KUKA KRL program: DrillingPart.src

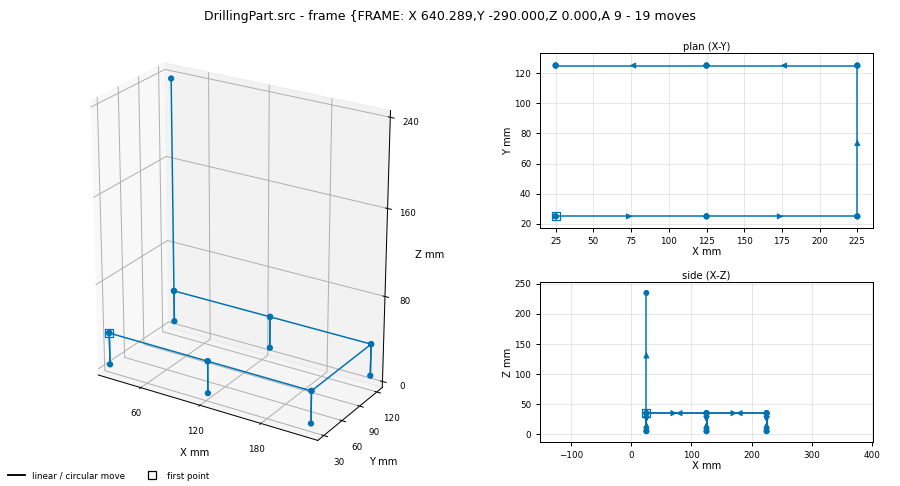
[picture p0: tool path of DrillingPart.src in frame {FRAME: X 640.289,Y -290.000,Z 0.000,A 9, 19 of 20 moves have a stored position in this frame; points joined in program order, loops and branches not executed]
&ACCESS RVP
&REL 1
&PARAM TEMPLATE = C:\KRC\Roboter\Template\vorgabe
&PARAM EDITMASK = *
DEF DrillingPart ( )
EXT BAS (BAS_COMMAND :IN,REAL :IN )


; GLOBAL INTERRUPT DECL 3 WHEN $STOPMESS==TRUE DO IR_STOPM ( )
; INTERRUPT ON 3

;FOLD Initialise and set default speed
BAS (#INITMOV,0)
BAS (#VEL_PTP,100)
BAS (#ACC_PTP,20)
$VEL.CP=0.2
BAS (#TOOL,0)
BAS (#BASE,0)
;ENDFOLD

;;FOLD STARTPOS
;$BWDSTART = FALSE
;PDAT_ACT = PDEFAULT
;BAS(#PTP_DAT)
;FDAT_ACT = {TOOL_NO 0,BASE_NO 0,IPO_FRAME #BASE}
;BAS(#FRAMES)
;;ENDFOLD

$ADVANCE = 5

;FOLD ---- Quickly skip BCO ----
; PTP $AXIS_ACT
;ENDFOLD

;FOLD ---- GO HOME ----
; PTP {A1 0.000, A2 -90.000, A3 90.000, A4 0.000, A5 0.000, A6 0.000, E1 0, E2 0, E3 0, E4 0, E5 0, E6 0}
;ENDFOLD


; Program generated by VerticalBot Studio for KUKA KR 10 R900 sixx on 25/10/2026 12:00:00
; Using nominal kinematics.
; ---- Setting reference (Base) ----
; BASE_DATA[1] = {FRAME: X 640.289,Y -290.000,Z 0.000,A 90.000,B 0.000,C 0.000}
$BASE = {FRAME: X 640.289,Y -290.000,Z 0.000,A 90.000,B 0.000,C 0.000}
; $BASE = BASE_DATA[1]
; --------------------------
; ---- Setting tool (TCP) ----
$TOOL = {FRAME: X 116.058,Y 0.000,Z 219.481,A 0.000,B 60.000,C 0.000}
; --------------------------
PTP {A1 40.16630,A2 -71.39490,A3 131.33300,A4 60.01490,A5 -40.15900,A6 -30.06660}
LIN {X 25.000,Y 25.000,Z 35.000,A 90.000,B 0.000,C -180.000}
LIN {X 25.000,Y 25.000,Z 5.000,A 90.000,B 0.000,C -180.000}
LIN {X 25.000,Y 25.000,Z 35.000,A 90.000,B 0.000,C -180.000}
LIN {X 125.000,Y 25.000,Z 35.000,A 90.000,B 0.000,C -180.000}
LIN {X 125.000,Y 25.000,Z 5.000,A 90.000,B 0.000,C -180.000}
LIN {X 125.000,Y 25.000,Z 35.000,A 90.000,B 0.000,C -180.000}
LIN {X 225.000,Y 25.000,Z 35.000,A 90.000,B 0.000,C -180.000}
LIN {X 225.000,Y 25.000,Z 5.000,A 90.000,B 0.000,C -180.000}
LIN {X 225.000,Y 25.000,Z 35.000,A 90.000,B 0.000,C -180.000}
LIN {X 225.000,Y 125.000,Z 35.000,A 90.000,B 0.000,C -180.000}
LIN {X 225.000,Y 125.000,Z 5.000,A 90.000,B 0.000,C -180.000}
LIN {X 225.000,Y 125.000,Z 35.000,A 90.000,B 0.000,C -180.000}
LIN {X 125.000,Y 125.000,Z 35.000,A 90.000,B 0.000,C -180.000}
LIN {X 125.000,Y 125.000,Z 5.000,A 90.000,B 0.000,C -180.000}
LIN {X 125.000,Y 125.000,Z 35.000,A 90.000,B 0.000,C -180.000}
LIN {X 25.000,Y 125.000,Z 35.000,A 90.000,B 0.000,C -180.000}
LIN {X 25.000,Y 125.000,Z 5.000,A 90.000,B 0.000,C -180.000}
LIN {X 25.000,Y 125.000,Z 35.000,A 90.000,B 0.000,C -180.000}
LIN {X 25.000,Y 125.000,Z 235.000,A 90.000,B 0.000,C -180.000}
END
